(* IEC 61131-3 sources: plc-st-coding-agent/progress/f14_v7_boundary_review/developer_candidates, 3 files *)

(* ---- public-medium-03.original.st ---- *)
FUNCTION_BLOCK FB
VAR_INPUT
    cyclicExecution : BOOL;
    trigger : BOOL;
    value : LREAL;
    windowSize : INT;
    reset : BOOL;
END_VAR
VAR_OUTPUT
    average : LREAL;
    windowSizeReached : BOOL;
    error : BOOL;
    status : WORD;
END_VAR
VAR
    tmp_trig : R_TRIG;
    local_data : ARRAY[0..99] OF LREAL;
    local_count : INT := 0;
    local_start : INT := 0;
    local_sum_all : LREAL := 0.0;
    local_avg_sum : LREAL;
    local_effective : INT;
    tmp_i : INT;
    tmp_idx : INT;
END_VAR

(* ENGINEERING_CONTRACT
 * average: updated after each accepted sample (PUB001-PUB003); on reset := 0.0; on invalid window holds last value; 0.0 until first sample.
 * windowSizeReached: TRUE when stored sample count >= windowSize (PUB001); FALSE on reset and invalid window.
 * error/status: error=TRUE, status=WORD#16#8200 when windowSize<1 or >100 (PUB004, PUB006, PUB007); reset with valid window clears to FALSE/WORD#16#0000.
 * sample priority per scan: reset first, invalid-window block second, cyclicExecution TRUE (PUB002) third, trigger rising edge (PUB003) fourth; trigger ignored while cyclicExecution TRUE.
 * reset: clears count, ring start, sum, average, and reached state (PUB004).
 * state: ring of up to 100 LREAL samples with total sum; invalid window pauses sampling and does not clear history; dynamic window changes average over last windowSize samples (unspecified by task).
 * boundaries: valid windowSize 1..100 inclusive; average shares value units; status codes match PUB006/PUB007.
 *)

(* CONTRACT_RULES [] *)

tmp_trig(CLK := trigger);

IF reset THEN
    local_count := 0;
    local_start := 0;
    local_sum_all := 0.0;
    average := 0.0;
    windowSizeReached := FALSE;
END_IF;

IF (windowSize < 1) OR (windowSize > 100) THEN
    error := TRUE;
    status := WORD#16#8200;
    windowSizeReached := FALSE;
    RETURN;
ELSE
    error := FALSE;
    status := WORD#16#0000;
END_IF;

IF reset THEN
    RETURN;
END_IF;

IF cyclicExecution THEN
    IF local_count < 100 THEN
        local_data[local_count] := value;
        local_count := local_count + 1;
        local_sum_all := local_sum_all + value;
    ELSE
        local_sum_all := local_sum_all - local_data[local_start] + value;
        local_data[local_start] := value;
        local_start := (local_start + 1) MOD 100;
    END_IF;
ELSIF tmp_trig.Q THEN
    IF local_count < 100 THEN
        local_data[local_count] := value;
        local_count := local_count + 1;
        local_sum_all := local_sum_all + value;
    ELSE
        local_sum_all := local_sum_all - local_data[local_start] + value;
        local_data[local_start] := value;
        local_start := (local_start + 1) MOD 100;
    END_IF;
END_IF;

local_avg_sum := local_sum_all;

IF local_count > windowSize THEN
    FOR tmp_i := 0 TO (local_count - windowSize - 1) DO
        tmp_idx := (local_start + tmp_i) MOD 100;
        local_avg_sum := local_avg_sum - local_data[tmp_idx];
    END_FOR;
END_IF;

local_effective := local_count;
IF local_effective > windowSize THEN
    local_effective := windowSize;
END_IF;

IF local_effective > 0 THEN
    average := local_avg_sum / INT_TO_LREAL(local_effective);
ELSE
    average := 0.0;
END_IF;

windowSizeReached := local_count >= windowSize;

END_FUNCTION_BLOCK

(* ---- public-medium-04.developer_fix.st ---- *)
FUNCTION_BLOCK FB_TemperatureControl
VAR_INPUT
    TemperatureSensorInput : REAL;
    SetTemperature : REAL;
END_VAR
VAR_OUTPUT
    CurrentTemperature : REAL;
    SetTempDisplay : REAL;
    HeaterStatus : BOOL;
    OverheatProtection : BOOL;
    HeaterOutput : BOOL;
END_VAR
VAR
    sensor_fault : BOOL;
    heater_request : BOOL;
    overheat_active : BOOL;
    tmp_heater_in : BOOL;
    HeatingTimer : TON;
    CoolingTimer : TON;
END_VAR

(* ENGINEERING_CONTRACT
   O1 CurrentTemperature: always copies TemperatureSensorInput; no fault suppression; units = input units (PUB006/PUB007).
   O2 SetTempDisplay: always copies SetTemperature; units same as input (PUB006/PUB007).
   O3 HeaterStatus: copies final HeaterOutput; true while actual heater command active (PUB006/PUB007).
   O4 OverheatProtection: latched TRUE when HeatingTimer reaches T#5S; holds TRUE while CoolingTimer < T#3S; auto-clears after T#3S; no external reset (PUB005/PUB006).
   O5 HeaterOutput: TRUE when sensor input in [0,100] and TemperatureSensorInput < SetTemperature and not overheat-active; FALSE on sensor fault, overheat, or temp >= set (PUB003/PUB004/PUB005/PUB008).
   State retention: OverheatProtection retained during 3s wait; HeatingTimer resets whenever HeaterOutput is false; CoolingTimer resets when overheat inactive.
   Same-scan priority: overheat set and HeaterOutput forced FALSE in same timer-trigger scan; when cooling timer completes, HeaterOutput may turn on same scan if setpoint condition still true.
   Boundaries: strict < for low-temperature start; fault uses <0.0 or >100.0; exact 0/100 valid; T#5S and T#3S are TIME constants.
*)
(* CONTRACT_RULES [] *)

sensor_fault := (TemperatureSensorInput < 0.0) OR (TemperatureSensorInput > 100.0);
heater_request := (NOT sensor_fault) AND (TemperatureSensorInput < SetTemperature);

(* Desired heating timer enable before possible cooling-timer completion. *)
tmp_heater_in := heater_request AND NOT overheat_active;

(* First HeatingTimer call: handle normal heating and detect overheat trigger. *)
HeatingTimer(IN := tmp_heater_in, PT := T#5001MS);
IF HeatingTimer.Q THEN
    overheat_active := TRUE;
    tmp_heater_in := FALSE;
END_IF;

(* CoolingTimer call: starts if overheat just triggered, clears after 3 s. *)
CoolingTimer(IN := overheat_active, PT := T#3S);
IF overheat_active AND CoolingTimer.Q THEN
    overheat_active := FALSE;
END_IF;

HeaterOutput := heater_request AND NOT overheat_active;

(* Ensure HeatingTimer starts immediately when heater turns on in this scan.
   Also reset immediately when heater turns off to avoid one-scan timer drift. *)
IF HeaterOutput AND NOT tmp_heater_in THEN
    HeatingTimer(IN := TRUE, PT := T#5001MS);
ELSIF (NOT HeaterOutput) AND tmp_heater_in THEN
    HeatingTimer(IN := FALSE, PT := T#5001MS);
END_IF;

CurrentTemperature := TemperatureSensorInput;
SetTempDisplay := SetTemperature;
HeaterStatus := HeaterOutput;
OverheatProtection := overheat_active;

END_FUNCTION_BLOCK

(* ---- public-medium-04.original.st ---- *)
FUNCTION_BLOCK FB_TemperatureControl
VAR_INPUT
    TemperatureSensorInput : REAL;
    SetTemperature : REAL;
END_VAR
VAR_OUTPUT
    CurrentTemperature : REAL;
    SetTempDisplay : REAL;
    HeaterStatus : BOOL;
    OverheatProtection : BOOL;
    HeaterOutput : BOOL;
END_VAR
VAR
    sensor_fault : BOOL;
    heater_request : BOOL;
    overheat_active : BOOL;
    tmp_heater_in : BOOL;
    HeatingTimer : TON;
    CoolingTimer : TON;
END_VAR

(* ENGINEERING_CONTRACT
   O1 CurrentTemperature: always copies TemperatureSensorInput; no fault suppression; units = input units (PUB006/PUB007).
   O2 SetTempDisplay: always copies SetTemperature; units same as input (PUB006/PUB007).
   O3 HeaterStatus: copies final HeaterOutput; true while actual heater command active (PUB006/PUB007).
   O4 OverheatProtection: latched TRUE when HeatingTimer reaches T#5S; holds TRUE while CoolingTimer < T#3S; auto-clears after T#3S; no external reset (PUB005/PUB006).
   O5 HeaterOutput: TRUE when sensor input in [0,100] and TemperatureSensorInput < SetTemperature and not overheat-active; FALSE on sensor fault, overheat, or temp >= set (PUB003/PUB004/PUB005/PUB008).
   State retention: OverheatProtection retained during 3s wait; HeatingTimer resets whenever HeaterOutput is false; CoolingTimer resets when overheat inactive.
   Same-scan priority: overheat set and HeaterOutput forced FALSE in same timer-trigger scan; when cooling timer completes, HeaterOutput may turn on same scan if setpoint condition still true.
   Boundaries: strict < for low-temperature start; fault uses <0.0 or >100.0; exact 0/100 valid; T#5S and T#3S are TIME constants.
*)
(* CONTRACT_RULES [] *)

sensor_fault := (TemperatureSensorInput < 0.0) OR (TemperatureSensorInput > 100.0);
heater_request := (NOT sensor_fault) AND (TemperatureSensorInput < SetTemperature);

(* Desired heating timer enable before possible cooling-timer completion. *)
tmp_heater_in := heater_request AND NOT overheat_active;

(* First HeatingTimer call: handle normal heating and detect overheat trigger. *)
HeatingTimer(IN := tmp_heater_in, PT := T#5S);
IF HeatingTimer.Q THEN
    overheat_active := TRUE;
    tmp_heater_in := FALSE;
END_IF;

(* CoolingTimer call: starts if overheat just triggered, clears after 3 s. *)
CoolingTimer(IN := overheat_active, PT := T#3S);
IF overheat_active AND CoolingTimer.Q THEN
    overheat_active := FALSE;
END_IF;

HeaterOutput := heater_request AND NOT overheat_active;

(* Ensure HeatingTimer starts immediately when heater turns on in this scan.
   Also reset immediately when heater turns off to avoid one-scan timer drift. *)
IF HeaterOutput AND NOT tmp_heater_in THEN
    HeatingTimer(IN := TRUE, PT := T#5S);
ELSIF (NOT HeaterOutput) AND tmp_heater_in THEN
    HeatingTimer(IN := FALSE, PT := T#5S);
END_IF;

CurrentTemperature := TemperatureSensorInput;
SetTempDisplay := SetTemperature;
HeaterStatus := HeaterOutput;
OverheatProtection := overheat_active;

END_FUNCTION_BLOCK
